(* IEC 61131-3 sources: st2fb/tests/fixtures/ecc/real_machines, 4 files *)

(* ---- fr1_linear_no_return.st ---- *)
FUNCTION_BLOCK LINEAR_START
VAR_INPUT GO : BOOL; READY : BOOL; END_VAR
VAR_OUTPUT STP : INT; CHARGING : BOOL; RUNNING : BOOL; END_VAR
  CHARGING := FALSE;
  CASE STP OF
    0: IF GO THEN STP := 1; END_IF;
    1: CHARGING := TRUE; IF READY THEN STP := 2; END_IF;
    2: RUNNING := TRUE;
  END_CASE;
END_FUNCTION_BLOCK

(* ---- fr2_retry_counter_guards.st ---- *)
FUNCTION_BLOCK RETRY_SM
VAR_INPUT GO : BOOL; OK : BOOL; RESET : BOOL; END_VAR
VAR_OUTPUT TRYING : BOOL; LOCKED : BOOL; TRIES : INT; END_VAR
VAR POS : INT; END_VAR
  TRYING := FALSE;
  CASE POS OF
    0: TRIES := 0; IF GO THEN POS := 1; END_IF;
    1: TRYING := TRUE;
       IF OK THEN POS := 0;
       ELSIF TRIES = 2 THEN LOCKED := TRUE; POS := 2;
       ELSE TRIES := TRIES + 1; END_IF;
    2: IF RESET THEN LOCKED := FALSE; POS := 0; END_IF;
  END_CASE;
END_FUNCTION_BLOCK

(* ---- fr3_hysteresis_integer.st ---- *)
FUNCTION_BLOCK HYST_SM
VAR_INPUT RAW : INT; END_VAR
VAR_OUTPUT PUMP : BOOL; FILTERED : INT; STARTS : INT; END_VAR
  IF PUMP THEN
    IF FILTERED < 5 THEN PUMP := FALSE; END_IF;
  ELSE
    IF FILTERED > 10 THEN PUMP := TRUE; STARTS := STARTS + 1; END_IF;
  END_IF;
  FILTERED := (FILTERED + RAW) / 2;
END_FUNCTION_BLOCK

(* ---- fr4_shared_mode_branch.st ---- *)
FUNCTION_BLOCK MODE_SM
VAR_INPUT GO : BOOL; SET_MODE : INT; END_VAR
VAR_OUTPUT ACTIVE : BOOL; RATE : INT; END_VAR
VAR GAIN : INT; END_VAR
  IF SET_MODE <> 0 THEN GAIN := SET_MODE; END_IF;
  IF ACTIVE THEN
    CASE GAIN OF 1: RATE := RATE + 1; 2: RATE := RATE + 2; END_CASE;
    IF NOT GO THEN ACTIVE := FALSE; END_IF;
  ELSE
    CASE GAIN OF 1: RATE := 0; 2: RATE := 100; END_CASE;
    IF GO THEN ACTIVE := TRUE; END_IF;
  END_IF;
END_FUNCTION_BLOCK
